(* PLC project TBEN_L5_PLC11.project, CODESYS CODESYS V3.5 SP21 Patch 1 *)
(* stored: creationDateTime 2026-11-07T15:35:08.4592076, modificationDateTime 2026-11-07T15:09:07.4034196 *)

// Ghi REAL dạng Float32T big-endian
FUNCTION F_IolSetR32BE : BOOL
VAR_INPUT
    pBuf  : POINTER TO BYTE;
    uiOff : UINT;
    rVal  : REAL;
END_VAR
VAR
    pDw : POINTER TO DWORD;
END_VAR

            pDw := ADR(rVal);
F_IolSetR32BE := F_IolSetU32BE(pBuf, uiOff, pDw^);

          
END_FUNCTION
